FUNCTION_BLOCK FB_sweep
VAR
	// VALORI DI INIZIALIZZAZIONE
	rStartFreq	:	REAL;
	rEndFreq	:	REAL;
	rLength		:	REAL;
	rK			:	REAL;
	
	// TIMER
	fbTimer			:	FB_Timer(T#0S);
END_VAR

METHOD ComputeFrequency : REAL
VAR_INPUT
END_VAR
ComputeFrequency	:=	F_interpolateReal(
	rX_Old	:=	0,
	rX_New	:=	rLength,
	rY_Old	:=	rStartFreq,
	rY_New	:=	rEndFreq,
	rX		:=	fbTimer.ComputeElapsedSeconds()
	);
END_METHOD

METHOD Initialize : BOOL
VAR_INPUT
	rInputStartFrequency	:	REAL;
	rInputEndFrequency		:	REAL;
	rInputLength			:	REAL;
END_VAR
rStartFreq	:=	rInputStartFrequency;
rEndFreq	:=	rInputEndFrequency;
rLength		:=	rInputLength;
rK			:=	(rEndFreq - rStartFreq) / rLength;

fbTimer.ChangeTimer(F_seconds2Time(rLength));
END_METHOD

ACTION Start:
fbTimer.Reset();
END_ACTION

METHOD Step : REAL
VAR_INPUT
END_VAR
VAR
	rTime	:	REAL;
END_VAR
IF fbTimer.VerifySelfElapsed() THEN
	Step	:=	0;
ELSE
	rTime	:=	fbTimer.ComputeElapsedSeconds();
	Step	:=	SIN(CONSTANTS.PI * rTime * (2 * rStartFreq + rK * rTime));
END_IF
END_METHOD

END_FUNCTION_BLOCK

(* stored: Version 1.1.0.1, ProductVersion 3.1.4024.9
   POU FB_sweep: Id {59b05527-a81a-46c0-8027-d759f6a264f9}, SpecialFunc None
   Folder ACTIONs: Id {430fb45c-a939-46a0-9118-70ab8b1d3642}
   Folder METHODs: Id {5bc75862-e8d2-426f-9b88-9dc79260b55d}
   Method ComputeFrequency: Id {3e1a0425-0a5c-4887-ba37-1e1bfc692f05}
   Method Initialize: Id {4d178d43-3de9-4702-8bed-ac650e456d29}
   Action Start: Id {39be2f7c-ee33-4e4c-838b-79b47bf8f887}
   Method Step: Id {38c0a492-17f1-43cd-ad95-a22e148d11c4} *)
